// TIA Portal V20 export
TYPE "WT_IO_Handbedienung _DIG_UDT"
   STRUCT
      iBetriebsart : Int;   // 0=Auto / 1=Hand EIN / 2=Hand AUS
      iZustand : Int;   // 0=AUS / 1=EIN / 10=Hand AUS / 11=Hand EIN
      byReserve : Array[0..5] of Byte;
   END_STRUCT;
END_TYPE
